// TIA Portal V21 export
// export: Created 2026-11-07T17:04:59.2247211Z, ExportSetting WithDefaults, DisplayName Totally Integrated Automation Portal, DisplayVersion V21, DisplayName STEP 7 Professional, DisplayVersion V21, DisplayName STEP 7 Safety, DisplayVersion V21, DisplayName Tech WebApplication, DisplayVersion V21, DisplayName WinCC Basic/Comfort/Advanced, DisplayVersion V21, DisplayName WinCC Unified, DisplayVersion V21
TextList "TL_Mode"  ListRange=Decimal
  TextListEntry   EntryType=SingleValue, Text="-"
  TextListEntry   EntryType=SingleValue, From=1, To=1, Text="AUTOMATSKI"
  TextListEntry   EntryType=SingleValue, From=2, To=2, Text="POLUAUTOMATSKI"
  TextListEntry   EntryType=SingleValue, From=3, To=3, Text="RUČNO"
